Fanuc KAREL source: KC00033.KL

PROGRAM KC00033
%NOLOCKGROUP
VAR
  I: INTEGER
  J: INTEGER
  K: INTEGER
  R: REAL
  B: BOOLEAN
  S: STRING[80]
  T: STRING[80]
  P: PATH
  Q: PATH
  AI: ARRAY[8] OF INTEGER
  AB: ARRAY[244] OF BYTE
  JP: JOINTPOS
  AR: ARRAY[6] OF REAL
BEGIN
  SET_PERCH(JP,AR,I)
END KC00033
